(* Rows filled in from the belt end down to where the entering rows have got to, a few per cycle. *)
un_FilledNow := 0;
WHILE un_FilledNow < un_STRESS_FILL_ROWS
AND lr_BeltLength - (UINT_TO_LREAL(un_FillRow) + 0.5) * lr_STRESS_PITCH > MIN(lr_BeltLength, lr_BeltPosition - lr_EntryStart) + lr_STRESS_PITCH / 2
AND DEMO_GlobalVar.DEMO_un_StressProducts > 0 DO
	m_LatchRow(lr_BeltLength - (UINT_TO_LREAL(un_FillRow) + 0.5) * lr_STRESS_PITCH);
	un_FillRow := un_FillRow + 1;
	un_FilledNow := un_FilledNow + 1;
END_WHILE

(* While switched off no rows enter: switched on again, the next one enters at the start, not rows behind it. *)
IF lr_BeltPosition - lr_NextRow > lr_STRESS_PITCH THEN
	lr_NextRow := lr_BeltPosition;
END_IF
IF lr_BeltPosition >= lr_NextRow AND DEMO_GlobalVar.DEMO_un_StressProducts > 0 THEN
	udn_RowFirstId[udn_RowCount MOD (VISU_GlobalConst_Param.VISU_un_MAX_PRODUCTS / 10 + 1)] := DEMO_GlobalVar.DEMO_udn_NextId;
	m_LatchRow(lr_STRESS_PITCH / 2 - (lr_BeltPosition - lr_NextRow));
	lr_NextRow := lr_NextRow + lr_STRESS_PITCH;
	(* One product of the row that entered half a belt ago is rejected: a state change on a full register. *)
	IF udn_RowCount >= un_Rows / 2 AND un_Rows > 1 THEN
		fb_StressBelt.m_SetProductState(
			vi_udn_Id := udn_RowFirstId[(udn_RowCount - un_Rows / 2) MOD (VISU_GlobalConst_Param.VISU_un_MAX_PRODUCTS / 10 + 1)]
				+ udn_RowCount MOD un_STRESS_LANES,
			vi_e_State := E_VisuProductState.REJECTED, vi_udn_ClientId := 0, vi_udn_MoverId := 0, vi_udn_FingerId := 0);
	END_IF
	udn_RowCount := udn_RowCount + 1;
END_IF


(****************************************************************************************************)
(* HOUSEKEEPING                                                                                     *)
(****************************************************************************************************)
fb_StressBelt.m_RemoveProductsBeyond(lr_BeltLength + DEMO_GlobalConst.DEMO_lr_REMOVE_BEYOND_END);
un_Products := fb_StressBelt.m_ProductCount();

(****************************************************************************************************<br>
© Syntegon Group.<br>
All rights reserved, also regarding any disposal, exploitation, reproduction, editing, distribution,<br>
as well as in the event of applications for industrial property rights.<br>
*****************************************************************************************************<br>
DESCRIPTION:<br>
Latches one row of products across the stress belt, one per lane, vi_lr_X mm from its start, with ids from<br>
DEMO_GlobalVar.DEMO_udn_NextId.<br>
*****************************************************************************************************<br>
OUTPUT VALUES:<br>
FALSE if a product did not fit into the register.<br>
****************************************************************************************************)
METHOD PRIVATE m_LatchRow : BOOL
VAR_INPUT
	vi_lr_X								: LREAL;	// [mm] along the belt from its start
END_VAR
VAR
	un_TempLane							: UINT;
	TempPose							: ST_VisuPlanarPose;
END_VAR
m_LatchRow := TRUE;
FOR un_TempLane := 0 TO un_STRESS_LANES - 1 DO
	TempPose.fX := vi_lr_X;
	TempPose.fY := lr_STRESS_Y + (UINT_TO_LREAL(un_TempLane) - UINT_TO_LREAL(un_STRESS_LANES - 1) / 2) * lr_STRESS_LANE_WIDTH;
	TempPose.fZ := DEMO_GlobalConst.DEMO_lr_BELT_Z;
	TempPose.fRz := 0;
	IF fb_StressBelt.m_LatchProduct(vi_udn_Id := DEMO_GlobalVar.DEMO_udn_NextId,
		vi_LatchPose := fb_StressBelt.m_McsToBelt(vi_Pose := TempPose),
		vi_udn_ProductType := 1, vi_lr_LatchBeltPosition := 0, vi_b_UseLatchBeltPosition := FALSE,
		vi_e_State := E_VisuProductState.DETECTED, vi_udn_ClientId := 0)
	THEN
		DEMO_GlobalVar.DEMO_udn_NextId := DEMO_GlobalVar.DEMO_udn_NextId + 1;
	ELSE
		m_LatchRow := FALSE;
	END_IF
END_FOR
END_METHOD

END_PROGRAM
